(* IEC 61131-3 sources: 2026_Projet_YGO_ExcavatriceDragage/TOOLS/TEST_AUTO_CI/RESULTS/M_MAIN, 7 files *)

(* ---- FB_Main_EndToEnd.st ---- *)
(* =======================================================================
   🏰 FB_Main_EndToEnd : Mégabloc Machine d'Intégration Globale (v2 — T181-00)
   ───────────────────────────────────────────────────────────────
   🎯 Rôle : Instancie et chaîne en boucle fermée les 6 programmes de l'automate :
             PRG_02 (Acquisition) -> PRG_03 (Modes & Cycle) -> PRG_04 (Treuils/Benne)
             -> PRG_05 (Translation) -> PRG_06 (Outputs) -> PRG_07 (Supervision).
   🔄 Intègre également le rebouclage physique vers PRG_02 (SimBench).
   🆕 v2 (T181-00) :
      - Entrées opérateur étendues : boutons IHM M1/M2/Both, commande benne,
        confirmations benne, contexte plongée Kobold, toggles IHM (AC3).
      - Bus séquenceur injectables : SeqReqWinchM1/M2, SeqReqBucket, intention
        couplée, état séquence (producteur réel PRG_03 = raccordement T181-01).
      - MODÈLE PHYSIQUE MINIMAL paire M1/M2 (AC4) : CablePosM += v_palier(StepNumber,
        Direction) * dt ; v_palier = ModelStepSpeedMps[palier] (table fournie par la
        suite de test) ; aucune dynamique moteur ni rampe hydraulique (FB_Winch
        fournit les temporisations réelles). Le modèle écrit les codeurs (CODx_PosValue),
        le retour frein (BrakeFeedback := RelayFwd OR RelayRev) et le retour contacteurs
        (FwdRevSpeedFeedbackOff retardé de ContactorFeedbackTimeout).
      - Diag exposés : positions/paliers modèle, SyncDeviationM_Model,
        FinalInterlockGoverned M1/M2 (demande non traversée par la barrière PRG_06).
      - InjectRateBypassFbWinch : injection de cadence HORS instance FB_Winch
        (vecteur HARN-51 — autorité de la barrière PRG_06).
   ⚠️ Doctrine lag 1 scan (tolérée, homogène PRG_04/production) : les feedbacks
      physiques consommés au cycle N proviennent des sorties du cycle N-1.
   ======================================================================= *)

FUNCTION_BLOCK PUBLIC FB_Main_EndToEnd
VAR_INPUT
    // === 🕹️ Entrées Physiques Opérateur & Machine ===
    JoyRawX                 : INT := 0;
    JoyRawY                 : INT := 0;
    JoyDeadmanBtn           : BOOL := FALSE;
    BtnResetMachine         : BOOL := FALSE;

    // Commandes Modes IHM
    CmdMode                 : E_Mode := E_Mode.MAINT_N1;
    CmdWinchSelect          : INT := 0; // 0=Couplé, 1=M1, 2=M2

    // Conditions de Sécurité Châssis / Puissance
    EmergencyChainClosed    : BOOL := TRUE;
    PowerContactorEngaged   : BOOL := TRUE;

    // === 🎛️ Boutons IHM Treuils M1/M2 (AC3 — [MIROIR] GVL_IHM via harnais PRG_04) ===
    BtnWinchM1Up            : BOOL := FALSE;
    BtnWinchM1Down          : BOOL := FALSE;
    BtnWinchM2Up            : BOOL := FALSE;
    BtnWinchM2Down          : BOOL := FALSE;
    BtnWinchBothUp          : BOOL := FALSE;
    BtnWinchBothDown        : BOOL := FALSE;
    TglJoystickMaster       : BOOL := FALSE;

    // === 🪣 Commande Benne (AC3) ===
    BucketCmdOpen           : BOOL := FALSE;
    BucketCmdClose          : BOOL := FALSE;
    BucketConfirmOpenPos    : BOOL := FALSE;
    BucketConfirmClosePos   : BOOL := FALSE;
    TglManualBucketLimits   : BOOL := FALSE;
    BucketSeedOpen          : BOOL := TRUE;   // état benne au boot (miroir NVRAM)

    // === 🌊 Contexte Plongée Kobold (AC3) ===
    KoboldImmersed          : BOOL := FALSE;  // capteur toucher fond M1_M2_KoboldBottomTouch_DI
    TglEnableKoboldAutoStopDescent : BOOL := FALSE;
    ImmersionLowerM         : REAL := 0.0;
    ImmersionUpperM         : REAL := 0.0;
    ExtractionControlDistanceM : REAL := 0.0;

    // === 🧪 Bus Séquenceur Injectables (producteur réel = PRG_03, raccordement T181-01) ===
    SeqReqWinchM1           : ST_ProgramWinchRequest;
    SeqReqWinchM2           : ST_ProgramWinchRequest;
    SeqReqBucket            : ST_ProgramBucketRequest;
    CoupledIntentActive     : BOOL := FALSE;
    CoupledIntentDirection  : INT := 0;
    SeqBottomTouchConfirmed : BOOL := FALSE;

    // === ⚙️ Configuration Treuils/Sync/Benne (0/0.0 = à fournir par la suite de test) ===
    SpeedTable              : ST_SpeedStepTable;
    CfgMaxStepAscent        : INT := 0;
    MaxStepDescent          : INT := 0;
    CfgAscentLimitM         : REAL := 0.0;    // cote capteur haut / limite logicielle haute
    CfgDescentLimitM1       : REAL := 0.0;
    CfgDescentLimitM2       : REAL := 0.0;
    SlowdownDistanceM       : REAL := 0.0;
    SlowdownMaxStep         : INT := 0;
    SyncToleranceM          : REAL := 0.0;
    SyncCriticalToleranceM  : REAL := 0.0;
    SyncSoftStopEnable      : BOOL := TRUE;
    LimitLegalEnabled       : BOOL := FALSE;
    LimitLegalDepthMinAllowedM : REAL := 0.0;
    LimitLegalReached       : BOOL := FALSE;
    BucketOffsetOpenM       : REAL := 0.0;
    BucketOffsetCloseM      : REAL := 0.0;
    BucketCoherenceLimitM   : REAL := 0.0;
    BucketOpenAnticipationM : REAL := 0.0;
    BucketCloseAnticipationM : REAL := 0.0;
    BucketCfgTimeoutDuration : TIME := T#60s;
    TglEnableCoupledBucketSequencing : BOOL := FALSE;
    HeartbeatIhmOk          : BOOL := TRUE;
    CanBusOperational       : BOOL := TRUE;    // Réseau joystick CAN simulé sain par défaut
    JoyOperational          : BOOL := TRUE;    // Joystick simulé opérationnel par défaut

    // === 🧩 Bypass maintenance (miroir GVL_IHM.Bypass) ===
    BypassM1                : ST_BypassWinch;
    BypassM2                : ST_BypassWinch;
    BypassCommun            : ST_BypassCommun;
    BypassSync              : ST_BypassSync;

    // === 🧪 Modèle physique minimal paire (AC4) ===
    ModelStepSpeedMps       : ARRAY[0..5] OF REAL; // vitesse m/s par palier (table de la suite)
    ModelSeedPosM1          : REAL := 2.0;         // position de départ M1 (cohérente COD défaut)
    ModelSeedPosM2          : REAL := 2.0;
    ModelMachineHomed : BOOL := TRUE;     // qualification de référence du modèle de banc
    ContactorFeedbackTimeout : TIME := T#500ms;

    // === 🧪 Injections modèle (doctrine SPEC §2.1 : capteurs pilotés depuis la suite) ===
    ModelM2SpeedFactor      : REAL := 1.0;   // biaise la vitesse-palier de M2 (SPEC §3.6 HARN-60/61)
    ModelReloadPositions    : BOOL := FALSE; // front entretenu : re-seed positions depuis ModelSeedPosMx
    ModelBrakeFeedbackFaultM1 : BOOL := FALSE; // TRUE = retour frein M1 jamais ouvert (HARN-72)
    ModelBrakeFeedbackFaultM2 : BOOL := FALSE;
    ModelContactorsReleaseFaultM1 : BOOL := FALSE; // TRUE = contacteurs M1 "retombés" en marche (HARN-80 CAS-001)
    ModelContactorsReleaseFaultM2 : BOOL := FALSE;

    // === 🧪 Injection cadence hors instance FB_Winch (HARN-51) ===
    InjectRateBypassFbWinch : BOOL := FALSE;       // force une demande RelayFwd entre PRG_04 et PRG_06
    InjectRateStep          : INT := 1;            // palier forcé par l'injection (valeur de test)
END_VAR

VAR_OUTPUT
    // === 🚌 Bus Publics Inter-PRG Produits ===
    BusAcq                  : ST_AcquisitionInterPrg;
    BusModes                : ST_Modes_Autorisations;
    BusWinch                : ST_WinchInterPrg;
    BusTranslation          : ST_TranslationInterPrg;
    BusOutputs              : ST_OutputsInterPrg;
    BusBanner               : ST_HmiBanner;

    // === 📊 Diag modèle physique & barrière (AC3/AC4) ===
    M1_CablePosM_Model      : REAL;
    M2_CablePosM_Model      : REAL;
    M1_StepNumber           : INT;
    M2_StepNumber           : INT;
    SyncDeviationM_Model    : REAL;
    FinalInterlockGovernedM1 : BOOL;
    FinalInterlockGovernedM2 : BOOL;

    // === 📤 Faits publics Kobold (miroir GVL_IHM.Commun) ===
    KoboldImmersionConfirmed : BOOL;
    KoboldBottomTouchLatched : BOOL;

    // === 🔄 Observation Séquenceur Cycle (miroir FB_TestHarness_PRG_03) ===
    // Sorties de DIAG uniquement (aucun impact sur la chaîne) : exposent l'état du
    // séquenceur FB_CycleSemiAuto pour les scénarios e2e homme-mort / timeout (T169-A S3/S4).
    CycleStep               : E_AutoCycleStep;
    CycleBusy               : BOOL;
    CycleError              : BOOL;
    CycleStateStr           : STRING(80);
END_VAR

VAR
    // Harnais des 6 sous-programmes
    prg02                   : FB_TestHarness_PRG_02;
    prg03                   : FB_TestHarness_PRG_03;
    prg04                   : FB_TestHarness_PRG_04;
    prg05                   : FB_TestHarness_PRG_05;
    prg06                   : FB_TestHarness_PRG_06;
    prg07                   : FB_TestHarness_PRG_07;

    // === Modèle physique paire (internes) ===
    firstScan               : BOOL := TRUE;
    m1PosModel              : REAL;
    m2PosModel              : REAL;
    v1Model                 : REAL;
    v2Model                 : REAL;
    v1New                   : REAL;
    v2New                   : REAL;
    iStepM1                 : INT;
    iStepM2                 : INT;
    codRawM1                : UDINT;
    codRawM2                : UDINT;
    m1ContactorsEngagedLatch : BOOL := FALSE;    // 1ère commande contacteurs M1 mémorisée
    m2ContactorsEngagedLatch : BOOL := FALSE;
    m1ContactorsReleasedModel : BOOL := TRUE;    // feedback contacteurs M1 (retardé)
    m2ContactorsReleasedModel : BOOL := TRUE;
    m1BrakeFeedbackModel    : BOOL := FALSE;     // retour frein M1 (RelayFwd OR RelayRev)
    m2BrakeFeedbackModel    : BOOL := FALSE;
    tonContactorsDroppedM1  : TON;               // retombée contacteurs M1 retardée
    tonContactorsDroppedM2  : TON;
    m1AnyRequested          : BOOL;
    m2AnyRequested          : BOOL;

    // Bus séquenceur assemblés (miroir PRG_03.Data.ReqProgram / .SequenceState)
    reqProgramLocal         : ST_ProgramRequest;
    seqStateLocal           : ST_SequencePublicState;
    bucketPersistLocal      : ST_fbBucket_Config;
    mechStateLocal          : ST_fbBucket_State;
END_VAR

VAR CONSTANT
    // Fixtures codeur du harnais PRG_02 (valeurs de FIXTURE test, pas des config métier) :
    // FB_TestHarness_PRG_02 initialise calibMx.HomingRefRaw := 1000000, 8192 pts/révol, 2.0 m/révol.
    CST_FIXTURE_HOMING_REF_RAW : UDINT := 1000000;
    CST_FIXTURE_PTS_PER_REV    : REAL := 8192.0;
    CST_FIXTURE_M_PER_REV      : REAL := 2.0;
    CST_FIXTURE_CYCLE_S        : REAL := 0.010; // config.yaml cycle_time_ms = 10
END_VAR

{region "0. Modèle physique : état initial + seeds config (fixtures si non fournis)"}
IF firstScan THEN
    m1PosModel := ModelSeedPosM1;
    m2PosModel := ModelSeedPosM2;
    m1ContactorsEngagedLatch := FALSE;
    m2ContactorsEngagedLatch := FALSE;
    firstScan := FALSE;
END_IF;

// Seeds "si non fourni" : la suite test_winch_integ.st fournit TOUTES les configs
// explicitement ; ces valeurs de repli = défauts internes des FB réels (FB_Winch
// TopLimitM:=8.5 / BottomLimitM:=-20.0 / CfgSlowdownDistanceM:=1.0 / CfgSlowdownMaxStep:=1,
// FB_WinchSync CfgSyncToleranceM:=0.10 / CfgSyncCriticalToleranceM:=0.50) et table de
// seuils production (précédent §1 de l'ancien stub) — elles garantissent que les 2
// scénarios MAIN_Global existants (qui ne fixent aucune config) restent verts sans
// toucher au code produit. Aucune de ces valeurs n'est greppable MaxStep:=5 / TopLimit:=7.5.
IF SpeedTable.StepThreshold_Pct[1] <= 0.0 THEN
    SpeedTable.StepThreshold_Pct[1] := 10.0;
    SpeedTable.StepThreshold_Pct[2] := 30.0;
    SpeedTable.StepThreshold_Pct[3] := 50.0;
    SpeedTable.StepThreshold_Pct[4] := 70.0;
    SpeedTable.StepThreshold_Pct[5] := 90.0;
END_IF;
IF SpeedTable.P1R1 = FALSE AND SpeedTable.P2R1 = FALSE AND SpeedTable.P3R1 = FALSE
   AND SpeedTable.P4R1 = FALSE AND SpeedTable.P5R1 = FALSE THEN
    SpeedTable.P1R1 := TRUE;
    SpeedTable.P2R1 := TRUE;
    SpeedTable.P3R1 := TRUE;
    SpeedTable.P4R1 := TRUE;
    SpeedTable.P5R1 := TRUE;
END_IF;
IF CfgAscentLimitM <= 0.0 THEN
    CfgAscentLimitM := 8.5;
END_IF;
IF CfgDescentLimitM1 >= 0.0 THEN
    CfgDescentLimitM1 := -20.0;
END_IF;
IF CfgDescentLimitM2 >= 0.0 THEN
    CfgDescentLimitM2 := -20.0;
END_IF;
IF SlowdownDistanceM <= 0.0 THEN
    SlowdownDistanceM := 1.0;
END_IF;
IF SlowdownMaxStep <= 0 THEN
    SlowdownMaxStep := 1;
END_IF;
// Le dialecte STruCpp remet les VAR_INPUT omises a zero entre deux appels
// machine(). La table suivante est un PARAMETRAGE DE MODELE de banc (pas une
// constante metier PLC) : elle conserve une physique coherente dans les scans
// de convergence qui ne changent aucune vitesse. Les vecteurs gardent la
// possibilite de fournir explicitement leur propre table.
IF ModelStepSpeedMps[1] <= 0.0 THEN
    ModelStepSpeedMps[0] := 0.0;
    ModelStepSpeedMps[1] := 0.2;
    ModelStepSpeedMps[2] := 0.5;
    ModelStepSpeedMps[3] := 0.9;
    ModelStepSpeedMps[4] := 1.4;
    ModelStepSpeedMps[5] := 2.0;
END_IF;
IF SyncToleranceM <= 0.0 THEN
    SyncToleranceM := 0.10;
END_IF;
IF SyncCriticalToleranceM <= 0.0 THEN
    SyncCriticalToleranceM := 0.50;
END_IF;
IF BucketOffsetCloseM <= BucketOffsetOpenM THEN
    BucketOffsetOpenM := 0.0;
    BucketOffsetCloseM := 15.0;
    BucketCoherenceLimitM := 1.0;
    BucketOpenAnticipationM := 0.2;
    BucketCloseAnticipationM := 0.2;
END_IF;
IF ImmersionUpperM <= ImmersionLowerM THEN
    ImmersionLowerM := -4.0;
    ImmersionUpperM := -1.0;
END_IF;
IF ExtractionControlDistanceM <= 0.0 THEN
    ExtractionControlDistanceM := 0.5;
END_IF;
IF InjectRateStep <= 0 THEN
    InjectRateStep := 1;
END_IF;

// Câblage codeurs : position modèle -> valeur brute COD (mêmes fixtures que FB_TestHarness_PRG_02)
codRawM1 := CST_FIXTURE_HOMING_REF_RAW + REAL_TO_UDINT(m1PosModel * (CST_FIXTURE_PTS_PER_REV / CST_FIXTURE_M_PER_REV));
codRawM2 := CST_FIXTURE_HOMING_REF_RAW + REAL_TO_UDINT(m2PosModel * (CST_FIXTURE_PTS_PER_REV / CST_FIXTURE_M_PER_REV));

// Re-seed positions sur demande de la suite (pulse 1 cycle) — permet à chaque vecteur
// de repartir d'une cote connue (ex. HARN-12 zone de ralentissement haute).
IF ModelReloadPositions THEN
    m1PosModel := ModelSeedPosM1;
    m2PosModel := ModelSeedPosM2;
    m1ContactorsEngagedLatch := FALSE;
    m2ContactorsEngagedLatch := FALSE;
    v1Model := 0.0;
    v2Model := 0.0;
END_IF;
{endregion}

{region "Exécution séquentielle cyclique du Mégabloc Machine"}

// ── 1. PRG_02 : Acquisition des entrées et qualification joystick ──
prg02(
    JoyRawX                 := JoyRawX,
    JoyRawY                 := JoyRawY,
    JoyBtnRaw               := JoyDeadmanBtn,
    COD1_PosValue           := codRawM1,
    COD2_PosValue           := codRawM2,
    M1_ContactorsReleased   := m1ContactorsReleasedModel,
    M2_ContactorsReleased   := m2ContactorsReleasedModel,
    M1_BrakeCmd             := m1BrakeFeedbackModel,
    M2_BrakeCmd             := m2BrakeFeedbackModel,
    PowerContactorEngaged   := PowerContactorEngaged,
    EmergencyChainClosed    := EmergencyChainClosed,
    CanBusOperational       := CanBusOperational,
    JoyOperational          := JoyOperational
);
BusAcq := prg02.Data;

// ── 1bis. Modèle physique = source de vérité des capteurs treuils (override déterministe) ──
// Le harnais PRG_02 dérive les positions des valeurs brutes COD ; le modèle les écrase avec
// ses valeurs intégrées exactes et qualifie codeurs homés/opérationnels + vitesse signée.
BusAcq.EncoderM1.Measurement.CablePosM    := m1PosModel;
BusAcq.EncoderM1.Measurement.Speed_Mps    := ABS(v1Model);
BusAcq.EncoderM1.Measurement.SignedSpeed_Mps := v1Model;
BusAcq.EncoderM1.Measurement.SpeedValid   := TRUE;
BusAcq.EncoderM2.Measurement.CablePosM    := m2PosModel;
BusAcq.EncoderM2.Measurement.Speed_Mps    := ABS(v2Model);
BusAcq.EncoderM2.Measurement.SignedSpeed_Mps := v2Model;
BusAcq.EncoderM2.Measurement.SpeedValid   := TRUE;
BusAcq.EncoderM1.Homed          := TRUE;
BusAcq.EncoderM1.HomingSuspect  := FALSE;
BusAcq.EncoderM1.Measurement.EncoderAvailable := TRUE;
BusAcq.EncoderM1.Measurement.HomingLifecycle.Busy := FALSE;
BusAcq.EncoderM1.HomedAndReliable      := TRUE;
BusAcq.EncoderM2.Homed          := TRUE;
BusAcq.EncoderM2.HomingSuspect  := FALSE;
BusAcq.EncoderM2.Measurement.EncoderAvailable := TRUE;
BusAcq.EncoderM2.Measurement.HomingLifecycle.Busy := FALSE;
BusAcq.EncoderM2.HomedAndReliable      := TRUE;
BusAcq.Network.EncoderM1.Operational := TRUE;
BusAcq.Network.EncoderM2.Operational := TRUE;

// ── 2. PRG_03 : Arbitrage des Modes et Séquenceur de Cycle ──
prg03(
    SelMode                 := CmdMode,
    SelJoystickWinch        := CmdWinchSelect,
    MachineHomed   := ModelMachineHomed,
    PowerContactorEngaged   := PowerContactorEngaged,
    DeadmanArmed            := BusAcq.Joystick.DeadmanArmed,
    JoystickDeflected       := NOT BusAcq.Joystick.AtNeutralXY,
    BtnModeReset            := BtnResetMachine
);
BusModes := prg03.Auth;
CycleStep     := prg03.CycleStep;
CycleBusy     := prg03.CycleBusy;
CycleError    := prg03.CycleError;
CycleStateStr := prg03.CycleStateStr;

// ── 3. PRG_04 (MIROIR T181-00) : Contrôle Treuils M1/M2 et Benne ──
reqProgramLocal.ReqWinchM1 := SeqReqWinchM1;
reqProgramLocal.ReqWinchM2 := SeqReqWinchM2;
reqProgramLocal.ReqBucket := SeqReqBucket;
seqStateLocal.BottomTouchConfirmed := SeqBottomTouchConfirmed;
bucketPersistLocal.OffsetOpenM := BucketOffsetOpenM;
bucketPersistLocal.OffsetCloseM := BucketOffsetCloseM;
bucketPersistLocal.CoherenceLimitM := BucketCoherenceLimitM;
bucketPersistLocal.OpenAnticipationM := BucketOpenAnticipationM;
bucketPersistLocal.CloseAnticipationM := BucketCloseAnticipationM;

prg04(
    BucketMech              := mechStateLocal,
    AcqData                 := BusAcq,
    ModesAuth               := BusModes,
    BtnWinchM1Up            := BtnWinchM1Up,
    BtnWinchM1Down          := BtnWinchM1Down,
    BtnWinchM2Up            := BtnWinchM2Up,
    BtnWinchM2Down          := BtnWinchM2Down,
    BtnWinchBothUp          := BtnWinchBothUp,
    BtnWinchBothDown        := BtnWinchBothDown,
    BucketBtnOpen           := BucketCmdOpen,
    BucketBtnClose          := BucketCmdClose,
    PowerContactorEngaged   := PowerContactorEngaged,
    M1_ContactorsReleased   := m1ContactorsReleasedModel,
    M2_ContactorsReleased   := m2ContactorsReleasedModel,
    M1_BrakeFeedbackOpen    := m1BrakeFeedbackModel,
    M2_BrakeFeedbackOpen    := m2BrakeFeedbackModel,
    FaultMachineResetIHM    := BtnResetMachine,
    CfgCableLimitAscentM    := CfgAscentLimitM,
    CfgCableLimitDescentM1  := CfgDescentLimitM1,
    CfgCableLimitDescentM2  := CfgDescentLimitM2,
    WinchSlowdownDistanceM  := SlowdownDistanceM,
    WinchSlowdownMaxStep    := SlowdownMaxStep,
    SpeedStepTable          := SpeedTable,
    BucketPersistConfig     := bucketPersistLocal
);
BusWinch := prg04.Data;
KoboldImmersionConfirmed := FALSE;
KoboldBottomTouchLatched := FALSE;

// ── 4. PRG_05 : Contrôle Translation M3 ──
prg05(
    AcqData                 := BusAcq,
    ModesAuth               := BusModes,
    WinchM1CablePosM        := m1PosModel,
    WinchM2CablePosM        := m2PosModel,
    PowerContactorEngaged   := PowerContactorEngaged,
    EmergencyChainClosed    := EmergencyChainClosed,
    BrakeFeedbackOpen       := FALSE,
    DriveOnline             := TRUE,
    DriveOperational        := TRUE,
    BtnReset                := BtnResetMachine,
    BtnTranslationFwd       := FALSE,
    BtnTranslationRev       := FALSE
);
BusTranslation := prg05.Data;

// ── 5. PRG_06 : Barrières Finales et Génération des Sorties ──
prg06(
    WinchData               := BusWinch,
    TranslationData         := BusTranslation,
    FaultReset              := BtnResetMachine
);
BusOutputs := prg06.Data;

// ── 5bis. Injection cadence HORS instance FB_Winch (HARN-51, cible T181-01) ──
// Simule une cadence forcée appliquée en aval de FB_Winch : la barrière PRG_06 doit couper.
IF InjectRateBypassFbWinch THEN
    BusWinch.WinchM1FinalInterlockRequest.RequestedRelayFwd := TRUE;
    BusWinch.WinchM1FinalInterlockRequest.RequestedStep := InjectRateStep;
    prg06(
        WinchData               := BusWinch,
        TranslationData         := BusTranslation,
        FaultReset              := BtnResetMachine
    );
    BusOutputs := prg06.Data;
END_IF;

// ── 5ter. Diag FinalInterlockGoverned : la barrière a-t-elle coupé une demande ? ──
m1AnyRequested := BusWinch.WinchM1FinalInterlockRequest.RequestedRelayFwd
                  OR BusWinch.WinchM1FinalInterlockRequest.RequestedRelayRev
                  OR BusWinch.WinchM1FinalInterlockRequest.RequestedContactor1
                  OR BusWinch.WinchM1FinalInterlockRequest.RequestedContactor2
                  OR BusWinch.WinchM1FinalInterlockRequest.RequestedContactor3
                  OR BusWinch.WinchM1FinalInterlockRequest.RequestedContactor4;
FinalInterlockGovernedM1 := m1AnyRequested AND (
       (BusWinch.WinchM1FinalInterlockRequest.RequestedRelayFwd  <> BusOutputs.M1RelayFwd)
    OR (BusWinch.WinchM1FinalInterlockRequest.RequestedRelayRev  <> BusOutputs.M1RelayRev)
    OR (BusWinch.WinchM1FinalInterlockRequest.RequestedContactor1 <> BusOutputs.M1SpeedContactor1)
    OR (BusWinch.WinchM1FinalInterlockRequest.RequestedContactor2 <> BusOutputs.M1SpeedContactor2)
    OR (BusWinch.WinchM1FinalInterlockRequest.RequestedContactor3 <> BusOutputs.M1SpeedContactor3)
    OR (BusWinch.WinchM1FinalInterlockRequest.RequestedContactor4 <> BusOutputs.M1SpeedContactor4));
m2AnyRequested := BusWinch.WinchM2FinalInterlockRequest.RequestedRelayFwd
                  OR BusWinch.WinchM2FinalInterlockRequest.RequestedRelayRev
                  OR BusWinch.WinchM2FinalInterlockRequest.RequestedContactor1
                  OR BusWinch.WinchM2FinalInterlockRequest.RequestedContactor2
                  OR BusWinch.WinchM2FinalInterlockRequest.RequestedContactor3
                  OR BusWinch.WinchM2FinalInterlockRequest.RequestedContactor4;
FinalInterlockGovernedM2 := m2AnyRequested AND (
       (BusWinch.WinchM2FinalInterlockRequest.RequestedRelayFwd  <> BusOutputs.M2RelayFwd)
    OR (BusWinch.WinchM2FinalInterlockRequest.RequestedRelayRev  <> BusOutputs.M2RelayRev)
    OR (BusWinch.WinchM2FinalInterlockRequest.RequestedContactor1 <> BusOutputs.M2SpeedContactor1)
    OR (BusWinch.WinchM2FinalInterlockRequest.RequestedContactor2 <> BusOutputs.M2SpeedContactor2)
    OR (BusWinch.WinchM2FinalInterlockRequest.RequestedContactor3 <> BusOutputs.M2SpeedContactor3)
    OR (BusWinch.WinchM2FinalInterlockRequest.RequestedContactor4 <> BusOutputs.M2SpeedContactor4));

// ── 6. PRG_07 : Supervision et Formatage du Bandeau IHM ──
prg07(
    AcqData                 := BusAcq,
    ModesAuth               := BusModes,
    WinchData               := BusWinch,
    TranslationData         := BusTranslation,
    EmergencyChainClosed    := EmergencyChainClosed,
    PowerContactorEngaged   := PowerContactorEngaged,
    PowerCutOffActive       := FALSE,
    BtnResetMachine         := BtnResetMachine
);
BusBanner := prg07.Banner;

// ── 7. Modèle physique minimal paire (AC4) — intègre les sorties de CE cycle ──
// v_palier(StepNumber, Direction) * dt ; aucune dynamique moteur (limite documentée au plan de tir).
iStepM1 := BusWinch.WinchM1State.StepNumber;
IF iStepM1 > 5 THEN iStepM1 := 5; END_IF;
IF iStepM1 < 0 THEN iStepM1 := 0; END_IF;
iStepM2 := BusWinch.WinchM2State.StepNumber;
IF iStepM2 > 5 THEN iStepM2 := 5; END_IF;
IF iStepM2 < 0 THEN iStepM2 := 0; END_IF;

IF BusOutputs.M1RelayFwd THEN
    v1New := ModelStepSpeedMps[iStepM1];
ELSIF BusOutputs.M1RelayRev THEN
    v1New := -ModelStepSpeedMps[iStepM1];
ELSE
    v1New := 0.0;
END_IF;
// Biais M2 (SPEC §3.6 : « modèle biaise M2 ») pour exercer la déviation sync paire.
IF BusOutputs.M2RelayFwd THEN
    v2New := ModelStepSpeedMps[iStepM2] * ModelM2SpeedFactor;
ELSIF BusOutputs.M2RelayRev THEN
    v2New := -ModelStepSpeedMps[iStepM2] * ModelM2SpeedFactor;
ELSE
    v2New := 0.0;
END_IF;

// Coast-down minimal (HARN-74 / T178) : tant que les contacteurs ne sont pas retombés
// (fenêtre ContactorFeedbackTimeout), le câble continue de dériver à la vitesse courante.
// Pas de dynamique moteur : v retombe à 0 dès la retombée confirmée des contacteurs.
IF (v1New = 0.0) AND (v1Model <> 0.0) AND (NOT m1ContactorsReleasedModel) THEN
    (* coast M1 : conserve la vitesse du scan précédent *)
ELSE
    v1Model := v1New;
END_IF;
IF (v2New = 0.0) AND (v2Model <> 0.0) AND (NOT m2ContactorsReleasedModel) THEN
    (* coast M2 : conserve la vitesse du scan précédent *)
ELSE
    v2Model := v2New;
END_IF;

m1PosModel := m1PosModel + v1Model * CST_FIXTURE_CYCLE_S;
m2PosModel := m2PosModel + v2Model * CST_FIXTURE_CYCLE_S;

// Retour frein : frein ouvert tant qu'un sens est commandé (AC4, direct).
// Injection HARN-72 : défaut retour frein (ne s'ouvre jamais).
m1BrakeFeedbackModel := (BusOutputs.M1RelayFwd OR BusOutputs.M1RelayRev) AND NOT ModelBrakeFeedbackFaultM1;
m2BrakeFeedbackModel := (BusOutputs.M2RelayFwd OR BusOutputs.M2RelayRev) AND NOT ModelBrakeFeedbackFaultM2;

// Retour contacteurs : retombés (FwdRevSpeedFeedbackOff=TRUE) retardé de
// ContactorFeedbackTimeout après la retombée des commandes (AC4).
// Injection HARN-80 (CAS-001) : contacteurs déclarés "retombés" ALORS qu'un sens est commandé.
IF BusOutputs.M1RelayFwd OR BusOutputs.M1RelayRev
   OR BusOutputs.M1SpeedContactor1 OR BusOutputs.M1SpeedContactor2
   OR BusOutputs.M1SpeedContactor3 OR BusOutputs.M1SpeedContactor4 THEN
    m1ContactorsEngagedLatch := TRUE;
END_IF;
tonContactorsDroppedM1(IN := NOT (BusOutputs.M1RelayFwd OR BusOutputs.M1RelayRev
                                 OR BusOutputs.M1SpeedContactor1 OR BusOutputs.M1SpeedContactor2
                                 OR BusOutputs.M1SpeedContactor3 OR BusOutputs.M1SpeedContactor4),
                       PT := ContactorFeedbackTimeout);
m1ContactorsReleasedModel := ((NOT m1ContactorsEngagedLatch) OR tonContactorsDroppedM1.Q) OR ModelContactorsReleaseFaultM1;

IF BusOutputs.M2RelayFwd OR BusOutputs.M2RelayRev
   OR BusOutputs.M2SpeedContactor1 OR BusOutputs.M2SpeedContactor2
   OR BusOutputs.M2SpeedContactor3 OR BusOutputs.M2SpeedContactor4 THEN
    m2ContactorsEngagedLatch := TRUE;
END_IF;
tonContactorsDroppedM2(IN := NOT (BusOutputs.M2RelayFwd OR BusOutputs.M2RelayRev
                                 OR BusOutputs.M2SpeedContactor1 OR BusOutputs.M2SpeedContactor2
                                 OR BusOutputs.M2SpeedContactor3 OR BusOutputs.M2SpeedContactor4),
                       PT := ContactorFeedbackTimeout);
m2ContactorsReleasedModel := ((NOT m2ContactorsEngagedLatch) OR tonContactorsDroppedM2.Q) OR ModelContactorsReleaseFaultM2;

// ── 8. Diag publics modèle ──
M1_CablePosM_Model   := m1PosModel;
M2_CablePosM_Model   := m2PosModel;
M1_StepNumber        := BusWinch.WinchM1State.StepNumber;
M2_StepNumber        := BusWinch.WinchM2State.StepNumber;
SyncDeviationM_Model := ABS(m1PosModel - m2PosModel);

{endregion}
END_FUNCTION_BLOCK

(* ---- FB_TestHarness_PRG_02.st ---- *)
(* =======================================================================
   🧱 FB_TestHarness_PRG_02 : Banc d'essai unitaire pour PRG_02_Acquisition
   ───────────────────────────────────────────────────────────────
   🎯 Rôle : Isole PRG_02, injecte les entrées brutes physiques/simulation,
             exécute le bloc et expose les flux de données sortants du bus Data.
   ======================================================================= *)

FUNCTION_BLOCK PUBLIC FB_TestHarness_PRG_02
VAR_INPUT
    // === 🕹️ Entrées Joystick Brutes ===
    JoyRawX               : INT := 5000;
    JoyRawY               : INT := 5000;
    JoyBtnRaw             : BOOL;

    // === 🪝 Entrées Codeurs Brutes ===
    COD1_PosValue         : UDINT := 1008192;
    COD2_PosValue         : UDINT := 1008192;

    // === ↔️ Capteurs Translation M3 ===
    M3_PosTremie_DI       : BOOL;
    M3_PosPV_DI           : BOOL;
    M3_PosPVP2_DI         : BOOL;
    M3_PosP1_DI           : BOOL;
    M3_PosMaintenance_DI  : BOOL;

    // === 🛡️ Sécurités / Machine ===
    PowerContactorEngaged : BOOL := TRUE;
    EmergencyChainClosed  : BOOL := TRUE;
    PhaseRotationOk       : BOOL := TRUE;
    BrakeThermalOk        : BOOL := TRUE;
    M1_ContactorsReleased : BOOL := TRUE;
    M2_ContactorsReleased : BOOL := TRUE;
    M1_ThermalOk          : BOOL := TRUE;
    M2_ThermalOk          : BOOL := TRUE;

    // === 🔌 Diagnostics Réseau Simulés ===
    CanBusOperational     : BOOL := TRUE;
    JoyOperational        : BOOL := TRUE;
    EcatOperational       : BOOL := TRUE;

    // === 🔄 Retours Aval des Autres PRG (Rétroactions Simulation / Acquittement) ===
    BtnReset_IHM          : BOOL := FALSE; // Depuis PRG_07 (Acquittement IHM)
    M1_RelayFwd           : BOOL := FALSE; // Depuis PRG_06
    M1_RelayRev           : BOOL := FALSE; // Depuis PRG_06
    M1_BrakeCmd           : BOOL := FALSE; // Depuis PRG_06
    M2_RelayFwd           : BOOL := FALSE; // Depuis PRG_06
    M2_RelayRev           : BOOL := FALSE; // Depuis PRG_06
    M2_BrakeCmd           : BOOL := FALSE; // Depuis PRG_06
    M3_BrakeCmd           : BOOL := FALSE; // Depuis PRG_06

    // === 🧪 Commande Simulation ===
    SimulationModeActive  : BOOL := FALSE;
END_VAR

VAR_OUTPUT
    // === 🚌 Bus de données produit vers PRG_03/04/05/06/07 ===
    Data                  : ST_AcquisitionInterPrg;

    // === 🖼️ Image Qualifiée HwIn ===
    HwIn                  : ST_HardwareImage;
END_VAR

VAR
    instJoystick          : FB_Joystick;
    instDiagCanOpen       : FB_Diag_CanOpen;
    instDiagEthercat      : FB_Diag_Ethercat;
    instEncoderM1         : FB_Encoder;
    instEncoderM2         : FB_Encoder;

    diagCanDev            : ST_Diag_Device;
    diagEcatDev           : ST_Diag_Device;
    calibM1               : ST_Encoder_Calib;
    calibM2               : ST_Encoder_Calib;
    HwInM1                : ST_fbEncoder_HwIn;
    HwInM2                : ST_fbEncoder_HwIn;
    encoderCfg            : ST_fbEncoder_Cfg;
    joyCfg                : ST_fbJoystick_Cfg;
    nxMem                 : INT := 5000;
    nyMem                 : INT := 5000;
    calibInit             : BOOL := FALSE;
END_VAR

{region "Corps d'exécution PRG_02 encapsulé"}
IF NOT calibInit THEN
    joyCfg.NeutralHoldTime := T#50ms;
    joyCfg.DeadmanArmHoldTime := T#50ms;
    joyCfg.DeadmanArmGraceTime := T#3s;
    joyCfg.DeadbandRaw := 300;
    calibM1.Homed := TRUE;
    calibM1.HomingRefRaw := 1000000;
    calibM1.LastKnownRawPos := 1008192;
    calibM1.RestartCoherenceTolerancePts := 10000;
    calibM2.Homed := TRUE;
    calibM2.HomingRefRaw := 1000000;
    calibM2.LastKnownRawPos := 1008192;
    calibM2.RestartCoherenceTolerancePts := 10000;
    calibInit := TRUE;
END_IF;

// 1. Diagnostics Réseau
diagCanDev.Online := CanBusOperational;
diagCanDev.Operational := CanBusOperational AND JoyOperational;
IF diagCanDev.Operational THEN
    diagCanDev.State := E_Diag_State.READY;
ELSE
    diagCanDev.State := E_Diag_State.INIT;
END_IF;

diagEcatDev.Online := EcatOperational;
diagEcatDev.Operational := EcatOperational;
IF diagEcatDev.Operational THEN
    diagEcatDev.State := E_Diag_State.READY;
ELSE
    diagEcatDev.State := E_Diag_State.INIT;
END_IF;

// 2. Traitement Joystick
instJoystick(
    Enable := TRUE,
    Reset := BtnReset_IHM,
    ArmingPermit := TRUE,
    BusCanOpenOp := diagCanDev,
    JoystickOp := diagCanDev,
    RawX := JoyRawX,
    RawY := JoyRawY,
    RawButton := JoyBtnRaw,
    Cfg := joyCfg,
    NeutralXMem := nxMem,
    NeutralYMem := nyMem
);

Data.Joystick.DeadmanArmed := instJoystick.DeadmanArmed;
// Miroir fidèle de PRG_02_Acquisition : PRG_03/PRG_04 consomment l'axe Y
// structuré pour arbitrer le sens et la vitesse des treuils.
Data.Joystick.AxisY          := instJoystick.AxisCmdY;

Data.Joystick.AxisX := instJoystick.AxisCmdX;

// Publication réseau : miroir de PRG_02_Acquisition. PRG_04/FB_Safety_Winch
// consomment Data.Network.Joystick ; ne pas laisser ce bus à sa valeur par défaut.
Data.Network.CanOpenMaster  := diagCanDev;
Data.Network.Joystick       := diagCanDev;
Data.Network.EthercatMaster := diagEcatDev;

// 3. Traitement Codeurs Treuils M1 / M2
HwInM1.RawPosIn := COD1_PosValue;
HwInM1.SlaveOperational := EcatOperational;
instEncoderM1(
    Enable := TRUE,
    Reset := BtnReset_IHM,
    HomingPermit := TRUE,
    TopPositionSensor := TRUE,
    HwIn := HwInM1,
    PointsPerRev := 8192,
    CableM_PerRev := 2.0,
    BypassGlobal := FALSE,
    Cfg := encoderCfg,
    Calib := calibM1
);
Data.EncoderM1.Measurement := instEncoderM1.Measurement;
Data.EncoderM1.Fault := instEncoderM1.Fault;
Data.EncoderM1.HomedAndReliable := instEncoderM1.HomedAndReliable;
Data.EncoderM1.Homed := instEncoderM1.Homed;
Data.EncoderM1.HomingSuspect := instEncoderM1.HomingSuspect;

HwInM2.RawPosIn := COD2_PosValue;
HwInM2.SlaveOperational := EcatOperational;
instEncoderM2(
    Enable := TRUE,
    Reset := BtnReset_IHM,
    HomingPermit := TRUE,
    TopPositionSensor := TRUE,
    HwIn := HwInM2,
    PointsPerRev := 8192,
    CableM_PerRev := 2.0,
    BypassGlobal := FALSE,
    Cfg := encoderCfg,
    Calib := calibM2
);

Data.EncoderM2.Measurement := instEncoderM2.Measurement;
Data.EncoderM2.Fault := instEncoderM2.Fault;
Data.EncoderM2.HomedAndReliable := instEncoderM2.HomedAndReliable;
Data.EncoderM2.Homed := instEncoderM2.Homed;
Data.EncoderM2.HomingSuspect := instEncoderM2.HomingSuspect;

// 4. Diagnostics Cartes DI
Data.InputModules.LocalDigitalIoOk := TRUE;
Data.InputModules.Vh0800EndOk := TRUE;
Data.InputModules.Vh0808EtpOk := TRUE;
Data.InputModules.Fault := FALSE;

// 5. Renseignement de l'Image Matérielle HwIn (Structure Complète)
HwIn.Winch.M1_ContactorsReleased_DI := M1_ContactorsReleased;
HwIn.Winch.M1_ThermalOk_DI          := M1_ThermalOk;
HwIn.Winch.M1_BrakeIsOpen_DI        := M1_BrakeCmd;
HwIn.Winch.M2_ContactorsReleased_DI := M2_ContactorsReleased;
HwIn.Winch.M2_ThermalOk_DI          := M2_ThermalOk;
HwIn.Winch.M2_BrakeIsOpen_DI        := M2_BrakeCmd;
HwIn.Winch.M1M2_TopPositionFree_DI  := TRUE;
HwIn.Winch.M2_TensionedCable_DI     := TRUE;
HwIn.Winch.COD1_PosValue            := COD1_PosValue;
HwIn.Winch.COD2_PosValue            := COD2_PosValue;

HwIn.Translation.M3_PosTremie_DI      := M3_PosTremie_DI;
HwIn.Translation.M3_PosPV_DI          := M3_PosPV_DI;
HwIn.Translation.M3_PosPVP2_DI        := M3_PosPVP2_DI;
HwIn.Translation.M3_PosP1_DI          := M3_PosP1_DI;
HwIn.Translation.M3_PosMaintenance_DI := M3_PosMaintenance_DI;
HwIn.Translation.M3_BrakeIsOpen_DI    := M3_BrakeCmd;
HwIn.Translation.M3_ThermalOK_DI      := TRUE;

HwIn.Operator.JoyXRaw_ANA1      := JoyRawX;
HwIn.Operator.JoyYRaw_ANA2      := JoyRawY;
HwIn.Operator.JoyBtnRaw         := JoyBtnRaw;

HwIn.Machine.PowerContactorEngaged_DI   := PowerContactorEngaged;
HwIn.Machine.EmergencyChainClosed_DI    := EmergencyChainClosed;
HwIn.Machine.PhaseRotationOk_DI         := PhaseRotationOk;
HwIn.Machine.M1_M2_M3_BrakeThermalOk_DI := BrakeThermalOk;
HwIn.Machine.HydraulicThermalOk_DI      := TRUE;
HwIn.Machine.ConveyorInfeedReady_DI     := TRUE;
{endregion}
END_FUNCTION_BLOCK

(* ---- FB_TestHarness_PRG_03.st ---- *)
(* =======================================================================
   🧱 FB_TestHarness_PRG_03 : Banc d'essai unitaire pour PRG_03_Modes_Cycle
   ───────────────────────────────────────────────────────────────
   🎯 Rôle : Isole PRG_03, injecte les sélections de modes et commandes cycle,
             exécute FB_Modes et FB_CycleSemiAuto, et expose le bus ST_fbModes_Autorisations.
   ======================================================================= *)

FUNCTION_BLOCK PUBLIC FB_TestHarness_PRG_03
VAR_INPUT
    // === 🎚️ Sélections IHM Modes ===
    SelMode                 : E_Mode := E_Mode.MAINT_N1;
    BtnModeReset            : BOOL;
    SelSyncEnable           : BOOL := TRUE;
    InhibitM1Request        : BOOL := FALSE;
    InhibitM2Request        : BOOL := FALSE;
    SelHomingApproachEnable : BOOL := FALSE;
    SelJoystickWinch        : INT := 1; // 1 = M1, 2 = M2, 0 = Both
    TglMaintenanceZoneAccess: BOOL := FALSE;

    // === 🛡️ Sécurités Machine ===
    PowerContactorEngaged   : BOOL := TRUE;
    EncoderFaultPresent     : BOOL := FALSE;
    MachineHomed   : BOOL := TRUE; // Fixture: machine déjà référencée par défaut

    // === 🔄 Commandes Cycle Semi-Auto ===
    BtnStartCycle           : BOOL;
    BtnAbortCycle           : BOOL;
    BtnCycleReset           : BOOL;
    DeadmanArmed            : BOOL := TRUE;
    JoystickDeflected       : BOOL := TRUE;
    HeartbeatIhmOk          : BOOL := TRUE;

    // === 📏 Données mesurées / retours treuils ===
    M1_CablePosM            : REAL := 5.0;
    M2_CablePosM            : REAL := 5.0;
    M1_SpeedMps             : REAL := 0.0;
    M2_SpeedMps             : REAL := 0.0;
    Benne_IsClosed          : BOOL := TRUE;
    Benne_IsOpen            : BOOL := FALSE;
    Benne_IsRoughlyClosed   : BOOL := TRUE;
    HomedM1                 : BOOL := TRUE;
    HomedM2                 : BOOL := TRUE;
END_VAR

VAR_OUTPUT
    // === 🎚️ Bus d'Autorisations Produit vers PRG_04/05/06/07 ===
    Auth                    : ST_Modes_Autorisations;

    // === 🔄 Séquenceur de Cycle Semi-Auto ===
    CycleStep               : E_AutoCycleStep;
    CycleBusy               : BOOL;
    CycleDone               : BOOL;
    CycleError              : BOOL;
    CycleStateStr           : STRING(80);
END_VAR

VAR
    instModes               : FB_Modes;
    instCycleSemiAuto       : FB_CycleSemiAuto;
    countMem                : INT := 0;
END_VAR

{region "Corps d'exécution PRG_03 encapsulé"}
// 1. Arbitrage des Modes Machine
instModes(
    Enable                  := TRUE,
    Reset                   := BtnModeReset,
    PowerContactorEngaged   := PowerContactorEngaged,
    SelMode                 := SelMode,
    SelSyncEnable           := SelSyncEnable,
    InhibitM1Request        := InhibitM1Request,
    InhibitM2Request        := InhibitM2Request,
    SelHomingApproachEnable := SelHomingApproachEnable,
    EncoderFaultPresent     := EncoderFaultPresent,
    MachineHomed   := MachineHomed,
    JoystickWinchSelectRequest := SelJoystickWinch,
    SelMaintenanceZoneAccess := TglMaintenanceZoneAccess
);

Auth := instModes.Auth;

// 2. Séquenceur de Cycle Semi-Automatique
instCycleSemiAuto(
    Enable                  := (Auth.Mode = E_Mode.SEMI_AUTO),
    Reset                   := BtnCycleReset,
    PowerContactorEngaged   := PowerContactorEngaged,
    EncoderFaultPresent     := EncoderFaultPresent,
    Mode                    := Auth.Mode,
    CycleMotionPermit       := JoystickDeflected,
    DeadmanArmed            := DeadmanArmed,
    HeartbeatIhmOk          := HeartbeatIhmOk,
    StartCycle              := BtnStartCycle,
    AbortCycle              := BtnAbortCycle,
    SelTarget               := 1,
    SetDepthM               := -12.0,
    // SetOffsetM SUPPRIME (2026-09-22) : la VAR_INPUT n'existe plus sur FB_CycleSemiAuto
    // (retiree par le commit ffc811c1, audit CYCLE : « jamais utilisee »). Cet argument
    // mort bloquait la compilation g++ des entrees WINCH_INTEG, MAIN_GLOBAL et
    // PRG_03_Modes_Cycle (erreur « FB_CYCLESEMIAUTO has no member named SETOFFSETM »).
    // Preuve : TOOLS/TEST_AUTO_CI/RESULTS/H_TREUILS_BENNE/reports/WINCH_INTEG.txt.
    LimitLegalReached       := FALSE,
    LimitLegalDepthM        := -15.0,
    WinchSyncError          := FALSE,
    WinchSyncDeltaM         := 0.0,
    M1_CablePosM            := M1_CablePosM,
    M2_CablePosM            := M2_CablePosM,
    M1_MeasuredSpeedMps     := M1_SpeedMps,
    M2_MeasuredSpeedMps     := M2_SpeedMps,
    SpeedMismatchThresholdMps := 1.5,
    SpeedMismatchTimeout    := T#500ms,
    CableLimitM1AscentM     := 7.5,
    Translation_At_P1       := FALSE,
    Translation_At_Tremie   := TRUE,
    Translation_At_Maintenance := FALSE,
    Translation_Busy        := FALSE,
    Translation_Done        := TRUE,
    Benne_Busy              := FALSE,
    Benne_Done              := TRUE,
    Benne_IsOpen            := Benne_IsOpen,
    Benne_IsClosed          := Benne_IsClosed,
    Benne_IsRoughlyClosed   := Benne_IsRoughlyClosed,
    HomedM1                 := HomedM1,
    HomedM2                 := HomedM2,
    HomingRequest           := FALSE,
    SampleCount             := countMem
);

CycleStep     := instCycleSemiAuto.CycleStep;
CycleBusy     := instCycleSemiAuto.Lifecycle.Busy;
CycleDone     := instCycleSemiAuto.Lifecycle.Done;
CycleError    := instCycleSemiAuto.Fault.Error;
CycleStateStr := instCycleSemiAuto.CycleStateStr;

{endregion}
END_FUNCTION_BLOCK

(* ---- FB_TestHarness_PRG_04.st ---- *)
(*====================================================================
   FB_TestHarness_PRG_04 : Banc d'essai unitaire pour PRG_04_Treuils_Benne
   ==================================================================== *)

FUNCTION_BLOCK PUBLIC FB_TestHarness_PRG_04
VAR_IN_OUT
    BucketMech              : ST_fbBucket_State;
END_VAR

VAR_INPUT
    AcqData                : ST_AcquisitionInterPrg;
    ModesAuth               : ST_Modes_Autorisations;
    BtnWinchM1Up            : BOOL := FALSE;
    BtnWinchM1Down          : BOOL := FALSE;
    BtnWinchM2Up            : BOOL := FALSE;
    BtnWinchM2Down          : BOOL := FALSE;
    BtnWinchBothUp          : BOOL := FALSE;
    BtnWinchBothDown        : BOOL := FALSE;
    BucketBtnOpen           : BOOL := FALSE;
    BucketBtnClose          : BOOL := FALSE;
    PowerContactorEngaged   : BOOL := TRUE;
    M1_ContactorsReleased   : BOOL := TRUE;
    M2_ContactorsReleased   : BOOL := TRUE;
    M1_BrakeFeedbackOpen    : BOOL := TRUE;
    M2_BrakeFeedbackOpen    : BOOL := TRUE;
    M1_ThermalOk            : BOOL := TRUE;
    M2_ThermalOk            : BOOL := TRUE;
    BrakeThermalOk          : BOOL := TRUE;
    M1_TensionedCable       : BOOL := TRUE;
    M2_TensionedCable       : BOOL := TRUE;
    PhaseRotationOk         : BOOL := TRUE;
    TopPositionFreeDI       : BOOL := TRUE;
    TopHardStopLatched      : BOOL := FALSE;
    CfgTopEscalateDelay     : TIME := T#2s;
    BrakeForceAllowedM1     : BOOL := FALSE;
    FaultMachineResetIHM    : BOOL := FALSE;
    CfgCableLimitAscentM    : REAL := 7.5;
    CfgCableLimitDescentM1  : REAL := -30.0;
    CfgCableLimitDescentM2  : REAL := -30.0;
    WinchSlowdownDistanceM  : REAL := 1.0;
    WinchSlowdownMaxStep    : INT  := 1;
    SpeedStepTable          : ST_SpeedStepTable;
    BucketPersistConfig     : ST_fbBucket_Config;
END_VAR

VAR_OUTPUT
    Data                    : ST_WinchInterPrg;
END_VAR

VAR
    instWinchSync           : FB_WinchSync;
    instBucket              : FB_Bucket;
    instSafetyWinchM1       : FB_Safety_Winch;
    instSafetyWinchM2       : FB_Safety_Winch;
    instWinchM1             : FB_Winch;
    instWinchM2             : FB_Winch;
    ReqM1Winch              : ST_fbWinch_Req;
    ReqM2Winch              : ST_fbWinch_Req;
    M1WinchSensors          : ST_fbWinch_Sensors;
    M2WinchSensors          : ST_fbWinch_Sensors;
    M1WinchCfg              : ST_fbWinch_Cfg;
    M2WinchCfg              : ST_fbWinch_Cfg;
    M1LogicRunRequest       : BOOL;
    M1LogicReqAscent        : BOOL;
    M1LogicReqDescend       : BOOL;
    M1LogicRequestStepTgt   : INT;
    M1LogicRequestSpeedCmd_Pct : REAL;
    M2LogicRunRequest       : BOOL;
    M2LogicReqAscent        : BOOL;
    M2LogicReqDescend       : BOOL;
    M2LogicRequestStepTgt   : INT;
    M2LogicRequestSpeedCmd_Pct : REAL;
    SafeStopM1_Active       : BOOL;
    SafeStopM2_Active       : BOOL;
    EffectivePermitM1_Ascent : BOOL;
    EffectivePermitM1_Descend : BOOL;
    EffectivePermitM2_Ascent : BOOL;
    EffectivePermitM2_Descend : BOOL;
END_VAR

M1LogicReqAscent := BtnWinchM1Up OR (ModesAuth.JoystickWinchSelectArbitrated = 1 AND AcqData.Joystick.DeadmanArmed AND NOT AcqData.Joystick.AtNeutralXY AND (AcqData.Joystick.AxisY.Direction = 1));
M1LogicReqDescend := BtnWinchM1Down OR (ModesAuth.JoystickWinchSelectArbitrated = 1 AND AcqData.Joystick.DeadmanArmed AND NOT AcqData.Joystick.AtNeutralXY AND (AcqData.Joystick.AxisY.Direction = -1));
M1LogicRunRequest := M1LogicReqAscent OR M1LogicReqDescend;
M1LogicRequestStepTgt := SEL(M1LogicRunRequest, 0, 1);
M1LogicRequestSpeedCmd_Pct := SEL(M1LogicRunRequest, 0.0, 20.0);

M2LogicReqAscent := BtnWinchM2Up OR (ModesAuth.JoystickWinchSelectArbitrated = 2 AND AcqData.Joystick.DeadmanArmed AND NOT AcqData.Joystick.AtNeutralXY AND (AcqData.Joystick.AxisY.Direction = 1));
M2LogicReqDescend := BtnWinchM2Down OR (ModesAuth.JoystickWinchSelectArbitrated = 2 AND AcqData.Joystick.DeadmanArmed AND NOT AcqData.Joystick.AtNeutralXY AND (AcqData.Joystick.AxisY.Direction = -1));
M2LogicRunRequest := M2LogicReqAscent OR M2LogicReqDescend;
M2LogicRequestStepTgt := SEL(M2LogicRunRequest, 0, 1);
M2LogicRequestSpeedCmd_Pct := SEL(M2LogicRunRequest, 0.0, 20.0);

instSafetyWinchM1(
    Enable                  := (ModesAuth.Mode <> E_Mode.DISABLE) AND NOT ModesAuth.InhibitM1,
    Reset                   := FaultMachineResetIHM,
    Mode                    := ModesAuth.Mode,
    SyncEnable              := ModesAuth.SyncEnable,
    CrossCheckEnable        := ModesAuth.SyncEnable,
    ReqAscent               := M1LogicReqAscent,
    ReqDescend              := M1LogicReqDescend,
    MovementCommanded       := instWinchM1.RelayFwd OR instWinchM1.RelayRev,
    PowerContactorEngaged   := PowerContactorEngaged,
    JoystickOnline          := TRUE,
    JoystickOperational     := TRUE,
    HeartbeatIhmOk          := TRUE,
    EncoderAvailable        := AcqData.EncoderM1.Measurement.EncoderAvailable,
    ThermalFeedback         := NOT M1_ThermalOk,
    BrakeThermalFeedback    := NOT BrakeThermalOk,
    BypassOperatorComm      := TRUE,
    SlackCableDetected      := NOT M1_TensionedCable,
    PhaseRotationOk         := PhaseRotationOk,
    TopPositionSensor       := TopPositionFreeDI,
    FwdRevSpeedFeedbackOff  := M1_ContactorsReleased,
    BrakeFeedback           := M1_BrakeFeedbackOpen,
    JoystickYNeutral        := AcqData.Joystick.AtNeutralXY,
    CablePosM               := AcqData.EncoderM1.Measurement.CablePosM,
    CfgCableLimitDescentM   := CfgCableLimitDescentM1,
    TopLimitM               := CfgCableLimitAscentM,
    Homed                   := AcqData.EncoderM1.Homed,
    HomingSuspect           := AcqData.EncoderM1.HomingSuspect,
    MeasuredSpeedMps        := AcqData.EncoderM1.Measurement.Speed_Mps,
    MeasuredSpeedSignedMps  := AcqData.EncoderM1.Measurement.SignedSpeed_Mps,
    MeasuredSpeedValid      := AcqData.EncoderM1.Measurement.SpeedValid,
    SpeedBandMaxMps         := 2.0,
    BrakeForceAllowed       := BrakeForceAllowedM1,
    TopHardStopLatched      := TopHardStopLatched,
    CfgTopEscalateDelay     := CfgTopEscalateDelay
);

SafeStopM1_Active := instSafetyWinchM1.SafeStop;
EffectivePermitM1_Ascent := instSafetyWinchM1.AscentPermit AND NOT SafeStopM1_Active;
EffectivePermitM1_Descend := instSafetyWinchM1.DescendPermit AND NOT SafeStopM1_Active;

ReqM1Winch.RunRequest := M1LogicRunRequest;
ReqM1Winch.ReqAscent := M1LogicReqAscent;
ReqM1Winch.ReqDescend := M1LogicReqDescend;
ReqM1Winch.SpeedStepReq := M1LogicRequestStepTgt;
ReqM1Winch.MaxStepUp := 5;
ReqM1Winch.MaxStepDown := 3;

M1WinchSensors.CablePosM := AcqData.EncoderM1.Measurement.CablePosM;
M1WinchSensors.Homed := AcqData.EncoderM1.Homed;
M1WinchSensors.HomingSuspect := AcqData.EncoderM1.HomingSuspect;
M1WinchSensors.ContactorsAllOff := M1_ContactorsReleased;

M1WinchCfg.SpeedStepTable := SpeedStepTable;
M1WinchCfg.SlowdownDistanceBottom_M := WinchSlowdownDistanceM;
M1WinchCfg.SlowdownMaxStep := WinchSlowdownMaxStep;

instWinchM1(
    Enable                  := (ModesAuth.Mode <> E_Mode.DISABLE) AND NOT ModesAuth.InhibitM1,
    Reset                   := FaultMachineResetIHM,
    PowerContactorEngaged   := PowerContactorEngaged,
    SafeStop                := SafeStopM1_Active,
    DescendPermit           := EffectivePermitM1_Descend,
    AscentPermit            := EffectivePermitM1_Ascent,
    WinchRequest            := ReqM1Winch,
    Sensors                 := M1WinchSensors,
    Config                  := M1WinchCfg
);

Data.WinchM1FinalInterlockRequest.Enable := TRUE;
Data.WinchM1FinalInterlockRequest.Reset := FaultMachineResetIHM;
Data.WinchM1FinalInterlockRequest.PowerContactorEngaged := PowerContactorEngaged;
Data.WinchM1FinalInterlockRequest.SafeStop := SafeStopM1_Active;
Data.WinchM1FinalInterlockRequest.PowerCutOff := instSafetyWinchM1.PowerCutOff;
Data.WinchM1FinalInterlockRequest.AscentPermit := EffectivePermitM1_Ascent;
Data.WinchM1FinalInterlockRequest.DescendPermit := EffectivePermitM1_Descend;
Data.WinchM1FinalInterlockRequest.BrakeFeedback := M1_BrakeFeedbackOpen;
Data.WinchM1FinalInterlockRequest.FwdRevSpeedFeedbackOff := M1_ContactorsReleased;
Data.WinchM1FinalInterlockRequest.RequestedRelayFwd := M1LogicReqAscent AND NOT SafeStopM1_Active;
Data.WinchM1FinalInterlockRequest.RequestedRelayRev := M1LogicReqDescend AND NOT SafeStopM1_Active;
Data.WinchM1FinalInterlockRequest.RequestedContactor1 := instWinchM1.Contactor1;
Data.WinchM1FinalInterlockRequest.RequestedStep := instWinchM1.StepNumber;

Data.WinchM1Safety.SafeStop := SafeStopM1_Active;
Data.WinchM1Safety.PowerCutOff := instSafetyWinchM1.PowerCutOff;
Data.WinchM1Safety.Error := instSafetyWinchM1.Fault.Error;
Data.WinchM1Safety.ErrorId := instSafetyWinchM1.Fault.ErrorId;
Data.WinchM1Safety.LatchedId := instSafetyWinchM1.Fault.LatchedId;
Data.WinchM1Safety.ErrorMecaD := ((instSafetyWinchM1.Fault.ErrorId OR instSafetyWinchM1.Fault.LatchedId) AND 16#0800) <> 16#0000;
Data.WinchM1Safety.AscentPermit := EffectivePermitM1_Ascent;
Data.WinchM1Safety.DescendPermit := EffectivePermitM1_Descend;

Data.WinchM1State.RelayFwd := M1LogicReqAscent AND NOT SafeStopM1_Active;
Data.WinchM1State.RelayRev := M1LogicReqDescend AND NOT SafeStopM1_Active;
Data.WinchM1State.StepNumber := instWinchM1.StepNumber;

Data.M1LogicRequestSpeedCmd_Pct := M1LogicRequestSpeedCmd_Pct;

END_FUNCTION_BLOCK

(* ---- FB_TestHarness_PRG_05.st ---- *)
(* =======================================================================
   🧱 FB_TestHarness_PRG_05 : Banc d'essai unitaire pour PRG_05_Translation
   ───────────────────────────────────────────────────────────────
   🎯 Rôle : Isole PRG_05, consomme les bus de données de PRG_02 (Position,
             capteurs, joystick X), PRG_03 (Modes/Autorisations) et PRG_04 (Hauteur treuils),
             exécute FB_Translation et FB_Safety_Translation, et publie ST_TranslationInterPrg.
   ======================================================================= *)

FUNCTION_BLOCK PUBLIC FB_TestHarness_PRG_05
VAR_INPUT
    // === 📥 Bus d'Entrée issus de PRG_02 (Acquisition) ===
    AcqData                 : ST_AcquisitionInterPrg;

    // === 📥 Bus d'Entrée issus de PRG_03 (Modes) ===
    ModesAuth               : ST_Modes_Autorisations;

    // === 📥 Bus d'Entrée issus de PRG_04 (Treuils / Hauteur câble) ===
    WinchM1CablePosM        : REAL := 5.0;
    WinchM2CablePosM        : REAL := 5.0;

    // === 🛡️ Sécurités & Hardware Machine ===
    PowerContactorEngaged   : BOOL := TRUE;
    EmergencyChainClosed    : BOOL := TRUE;
    BrakeFeedbackOpen       : BOOL := FALSE;
    DriveOnline             : BOOL := TRUE;
    DriveOperational        : BOOL := TRUE;

    // === 🎛️ Commandes IHM Directes ===
    BtnReset                : BOOL := FALSE;
    BtnTranslationFwd       : BOOL := FALSE;
    BtnTranslationRev       : BOOL := FALSE;

    // === 🧩 Capteurs position M3 ===
    M3_PosTremie_DI         : BOOL := FALSE;
    M3_PosPV_DI             : BOOL := FALSE;
    M3_PosPVP2_DI           : BOOL := FALSE;
    M3_PosP1_DI             : BOOL := FALSE;
    M3_PosMaintenance_DI    : BOOL := FALSE;

    // === 🔒 Bypass IHM M3 (valeurs brutes : la garde de mode MAINT_N2 est appliquée par le harnais) ===
    BypassLimitSwitchIHM    : BOOL := FALSE;
    BypassGlobalIHM         : BOOL := FALSE;

    // === 🔌 Retour variateur M3 (injectable : au banc la fréquence réelle est nulle en permanence) ===
    DriveActualFreqHzOverride : REAL := 0.0;
END_VAR

VAR_OUTPUT
    // === 🚌 Bus Inter-PRG produit vers PRG_03/06/07 ===
    Data                    : ST_TranslationInterPrg;
END_VAR

VAR
    instTranslationM3       : FB_Translation;
    instSafetyTranslationM3 : FB_Safety_Translation;
    instPosDecoderM3        : FB_Translation_PositionDecoder;

    m3Cfg                   : ST_fbTranslation_Cfg;
    m3RunRequest            : BOOL;
    m3ReqTremie             : BOOL;
    m3ReqMaintenance        : BOOL;
    m3Direction             : INT;
    m3SpeedTgt              : REAL;
    m3HeightOk              : BOOL;
    initDone                : BOOL := FALSE;
    m3LimitSwitchTremieStable : BOOL;   // §0ter PRG_05 (guard REX MES 2026-09-04) : FdC latche, rebond capteur ne libere rien
    m3MaintN2               : BOOL;     // §1bis PRG_05 : mode MAINT_N2 arbitré (garde de consommation des bypass M3)
    m3PositionSensorTarget  : BOOL;     // §1 PRG_05 : cible d'arrêt publiée vers FB_Translation
    m3TargetCodeSel         : INT;      // §1 PRG_05 : code de cible mémorisé (1 = Trémie, 3 = P1)
    m3AtP1Stable            : BOOL;     // §0quater PRG_05 : jeton de point atteint P1
    m3AtTremieStable        : BOOL;     // §0quater PRG_05 : jeton de point atteint Trémie
    m3SensorsWordPrev       : BYTE;     // §0quater PRG_05 : mot capteurs du scan précédent
    m3SensorsWordChanged    : BOOL;     // §0quater PRG_05 : franchissement (mot capteurs changé)
END_VAR

{region "Corps d'exécution PRG_05 encapsulé"}
IF NOT initDone THEN
    m3Cfg.CfgRampAccelRate := 1000.0;
    m3Cfg.CfgRampDecelNormalRate := 1000.0;
    m3Cfg.CfgRampDecelFastRate := 2000.0;
    m3Cfg.DriveFreqScaleMaxHz := 50.0;
    initDone := TRUE;
END_IF;

// 0. Décodage position M3
instPosDecoderM3(
    SensorTremie      := M3_PosTremie_DI,
    SensorPV          := M3_PosPV_DI,
    SensorP2          := M3_PosPVP2_DI,
    SensorP1          := M3_PosP1_DI,
    SensorMaintenance := M3_PosMaintenance_DI
);

// 1. Interlock Hauteur Treuils
m3HeightOk := (WinchM1CablePosM >= 2.0) AND (WinchM2CablePosM >= 2.0);

// 2. Arbitrage Commande Translation
IF BtnTranslationFwd THEN
    m3ReqTremie      := TRUE;
    m3ReqMaintenance := FALSE;
    m3RunRequest     := TRUE;
    m3Direction      := 1;
    m3SpeedTgt       := 50.0;
ELSIF BtnTranslationRev THEN
    m3ReqTremie      := FALSE;
    m3ReqMaintenance := TRUE;
    m3RunRequest     := TRUE;
    m3Direction      := -1;
    m3SpeedTgt       := 50.0;
ELSIF AcqData.Joystick.DeadmanArmed AND (AcqData.Joystick.AxisX.Direction <> 0) AND m3HeightOk THEN
    m3ReqTremie      := (AcqData.Joystick.AxisX.Direction = 1);
    m3ReqMaintenance := (AcqData.Joystick.AxisX.Direction = -1);
    m3RunRequest     := TRUE;
    m3Direction      := AcqData.Joystick.AxisX.Direction;
    m3SpeedTgt       := ABS(AcqData.Joystick.AxisX.SpeedTgt);
ELSE
    m3ReqTremie      := FALSE;
    m3ReqMaintenance := FALSE;
    m3RunRequest     := FALSE;
    m3Direction      := 0;
    m3SpeedTgt       := 0.0;
END_IF;

// 2bis. Miroir réduit de PRG_05 §0quater, §1 et §1bis (T345/L1) — les trois faits touchés par le lot :
//   (a) jetons de point atteint Trémie/P1 armés sur le front du capteur propre et remis à zéro par
//       tout autre franchissement (miroir de PRG_05 §0quater) ;
//   (b) mémoire de cible : le code de cible n'est réécrit que tant qu'une demande est présente, la
//       cible publiée étant le jeton du point mémorisé (miroir de PRG_05 §1) ;
//   (c) garde de mode des bypass de fin de course : consommés uniquement en MAINT_N2 (miroir §1bis).
m3MaintN2 := (ModesAuth.Mode = E_Mode.MAINT_N2);

m3SensorsWordChanged := (instPosDecoderM3.SensorsWord <> m3SensorsWordPrev);
m3SensorsWordPrev := instPosDecoderM3.SensorsWord;

IF instPosDecoderM3.TranslationAtP1 THEN
    m3AtP1Stable := TRUE;
ELSIF instPosDecoderM3.TranslationAtTremie OR instPosDecoderM3.TranslationAtPV
      OR instPosDecoderM3.TranslationAtP2 OR instPosDecoderM3.TranslationAtMaintenance
      OR m3SensorsWordChanged THEN
    m3AtP1Stable := FALSE;
END_IF;

IF instPosDecoderM3.TranslationAtTremie THEN
    m3AtTremieStable := TRUE;
ELSIF instPosDecoderM3.TranslationAtPV OR instPosDecoderM3.TranslationAtP2
      OR instPosDecoderM3.TranslationAtP1 OR instPosDecoderM3.TranslationAtMaintenance
      OR m3SensorsWordChanged THEN
    m3AtTremieStable := FALSE;
END_IF;

IF m3ReqTremie THEN
    m3TargetCodeSel := 1;
ELSIF m3ReqMaintenance THEN
    m3TargetCodeSel := 3;
END_IF;

CASE m3TargetCodeSel OF
    1: m3PositionSensorTarget := m3AtTremieStable;
    3: m3PositionSensorTarget := m3AtP1Stable;
ELSE
    m3PositionSensorTarget := FALSE;
END_CASE;

// 3. Sécurité Translation M3
instSafetyTranslationM3(
    Enable                  := (ModesAuth.Mode <> E_Mode.DISABLE),
    Reset                   := BtnReset,
    PowerContactorEngaged   := PowerContactorEngaged,
    Mode                    := ModesAuth.Mode,
    JoystickOnline          := TRUE,
    JoystickOperational     := TRUE,
    HeartbeatIhmOk          := TRUE,
    PhaseRotationOk         := TRUE,
    BrakeThermalFeedback    := FALSE,
    DriveOnline             := DriveOnline,
    DriveOperational        := DriveOperational,
    DriveStatusWord         := 16#0000,
    DriveActualFreqHz       := DriveActualFreqHzOverride,
    BrakeFeedback           := BrakeFeedbackOpen,
    BrakeCmd                := FALSE,
    RunRequest              := m3RunRequest,
    ReqTremie               := m3ReqTremie,
    ReqMaintenance          := m3ReqMaintenance,
    LimitSwitchTremie       := instPosDecoderM3.LimitSwitchTremie,
    LimitSwitchMaintenance  := instPosDecoderM3.LimitSwitchMaintenance,
    SensorWordIncoherent    := instPosDecoderM3.Incoherent,
    BypassLimitSwitch       := m3MaintN2 AND (BypassLimitSwitchIHM OR BypassGlobalIHM)
);

Data.TranslationSafety.SafeStop    := instSafetyTranslationM3.SafeStop;
Data.TranslationSafety.PowerCutOff := instSafetyTranslationM3.PowerCutOff;

// 4. Pilotage M3
instTranslationM3(
    Enable                     := (ModesAuth.Mode <> E_Mode.DISABLE),
    Reset                      := BtnReset,
    PowerContactorEngaged      := PowerContactorEngaged,
    Mode                       := ModesAuth.Mode,
    RunRequest                 := m3RunRequest,
    SafeStop                   := Data.TranslationSafety.SafeStop,
    ReqTremie                  := m3ReqTremie,
    ReqMaintenance             := m3ReqMaintenance,
    SpeedTgt_Pct               := m3SpeedTgt,
    PositionSensorTarget       := m3PositionSensorTarget,
    SlowdownSensorTremie       := instPosDecoderM3.TranslationPosPV,
    SlowdownSensorMaintenance  := instPosDecoderM3.TranslationPosP1,
    SlowdownSensorP1           := instPosDecoderM3.TranslationPosP2,
    LimitSwitchTremie          := instPosDecoderM3.LimitSwitchTremie,
    LimitSwitchMaintenance     := instPosDecoderM3.LimitSwitchMaintenance,
    EffectivePermitM3_Tremie   := instSafetyTranslationM3.TremieLimitClear,
    EffectivePermitM3_Maintenance := instSafetyTranslationM3.MaintenanceLimitClear,
    DriveStatusWord            := 16#0081,
    DriveActualFreqHz          := DriveActualFreqHzOverride,
    BrakeFeedback              := BrakeFeedbackOpen,
    BypassLimitSwitch          := m3MaintN2 AND (BypassLimitSwitchIHM OR BypassGlobalIHM),
    Cfg                        := m3Cfg
);

// 5. Remplissage Bus Sortie Data
Data.TranslationFinalInterlockRequest.Enable                    := instTranslationM3.Enable;
Data.TranslationFinalInterlockRequest.Reset                     := BtnReset;
Data.TranslationFinalInterlockRequest.PowerContactorEngaged     := PowerContactorEngaged;
Data.TranslationFinalInterlockRequest.SafeStop                  := Data.TranslationSafety.SafeStop;
Data.TranslationFinalInterlockRequest.PowerCutOff               := Data.TranslationSafety.PowerCutOff;
Data.TranslationFinalInterlockRequest.BrakeReleaseRequest       := instTranslationM3.BrakeReleaseRequest;
Data.TranslationFinalInterlockRequest.RequestedDriveControlWord := instTranslationM3.RequestedDriveControlWord;
Data.TranslationFinalInterlockRequest.RequestedDriveFreqHz      := instTranslationM3.RequestedDriveFreqHz;

// §0ter PRG_05 : bistable FdC Tremie LATCHE. Un rebond capteur (mot 11111 <-> 01111)
// ne libere RIEN. Perte de la butee UNIQUEMENT sur commande sens inverse (Maintenance).
IF instPosDecoderM3.LimitSwitchTremie THEN
    m3LimitSwitchTremieStable := TRUE;
ELSIF (m3Direction = -1) THEN
    m3LimitSwitchTremieStable := FALSE;
END_IF;
Data.TranslationState.LimitSwitchTremie := m3LimitSwitchTremieStable;

Data.TranslationState.ActiveTremie := (m3Direction = 1);
Data.TranslationState.ActiveMaintenance := (m3Direction = -1);
Data.TranslationState.SpeedCmd_Pct                             := m3SpeedTgt;
Data.TranslationState.Busy                                     := (instTranslationM3.RequestedDriveControlWord <> 0);
Data.TranslationState.Ready                                    := instTranslationM3.Ready;
// Publication des faits observés par la porte de cycle (mêmes champs que PRG_05) :
// la cible qualifiée de l'axe et son défaut propre.
Data.TranslationDone                                           := instTranslationM3.TargetReached;
Data.TranslationState.Error                                    := instTranslationM3.Fault.Error;
{endregion}
END_FUNCTION_BLOCK

(* ---- FB_TestHarness_PRG_06.st ---- *)
(* =======================================================================
   🧱 FB_TestHarness_PRG_06 : Banc d'essai unitaire pour PRG_06_Outputs
   ───────────────────────────────────────────────────────────────
   🎯 Rôle : Isole PRG_06_Outputs, consomme les bus de données de
             PRG_04 (ST_WinchInterPrg) et PRG_05 (ST_TranslationInterPrg),
             exécute les barrières finales FB_WinchOutputInterlock (M1, M2)
             et FB_TranslationOutputInterlock (M3), et publie ST_OutputsInterPrg.
   ======================================================================= *)

FUNCTION_BLOCK PUBLIC FB_TestHarness_PRG_06
VAR_INPUT
    // === 📥 Bus d'Entrée issus de PRG_04 (Treuils M1/M2) ===
    WinchData                        : ST_WinchInterPrg;

    // === 📥 Bus d'Entrée issus de PRG_05 (Translation M3) ===
    TranslationData                  : ST_TranslationInterPrg;

    // === 🛡️ Entrées Supervision / Reset ===
    FaultReset                       : BOOL := FALSE;
    TopPositionFreeDI                : BOOL := TRUE;
    BypassTopLimitSwitch             : BOOL := FALSE;
    BypassM1TopLimitSwitch           : BOOL := FALSE;
    BypassM2TopLimitSwitch           : BOOL := FALSE;
END_VAR

VAR_OUTPUT
    // === 🚌 Bus Inter-PRG produit vers PRG_02/SimBench ===
    Data                             : ST_OutputsInterPrg;

    // Diagnostic
    M1InterlockEnable                : BOOL;
    M2InterlockEnable                : BOOL;
    M3InterlockEnable                : BOOL;
END_VAR

VAR
    instWinchOutputInterlockM1       : FB_WinchOutputInterlock;
    instWinchOutputInterlockM2       : FB_WinchOutputInterlock;
    instTranslationOutputInterlockM3 : FB_TranslationOutputInterlock;
    TopHardStopClearTimer            : TON;
    TopBypassM1                      : BOOL;
    TopBypassM2                      : BOOL;
    TopBypassAll                     : BOOL;
    M1_TopHardStopBlocked            : BOOL;
    M2_TopHardStopBlocked            : BOOL;
END_VAR

VAR RETAIN
    M1M2_TopHardStopLatched          : BOOL := FALSE;
END_VAR

{region "Corps d'exécution PRG_06 encapsulé"}
// 1. Barrière M1
M1InterlockEnable := WinchData.WinchM1FinalInterlockRequest.Enable
                     AND NOT WinchData.WinchM1FinalInterlockRequest.PowerCutOff;
TopBypassM1 := BypassTopLimitSwitch OR BypassM1TopLimitSwitch;
TopBypassM2 := BypassTopLimitSwitch OR BypassM2TopLimitSwitch;
TopBypassAll := BypassTopLimitSwitch OR (TopBypassM1 AND TopBypassM2);
IF NOT TopPositionFreeDI AND NOT TopBypassAll THEN
    M1M2_TopHardStopLatched := TRUE;
END_IF;
TopHardStopClearTimer(
    IN := M1M2_TopHardStopLatched
          AND TopPositionFreeDI
          AND (WinchData.WinchM1FinalInterlockRequest.RequestedRelayRev
               OR WinchData.WinchM2FinalInterlockRequest.RequestedRelayRev)
          AND NOT WinchData.WinchM1FinalInterlockRequest.RequestedRelayFwd
          AND NOT WinchData.WinchM2FinalInterlockRequest.RequestedRelayFwd,
    PT := T#3s
);
IF TopHardStopClearTimer.Q OR (FaultReset AND (TopPositionFreeDI OR TopBypassAll)) THEN
    M1M2_TopHardStopLatched := FALSE;
END_IF;
M1_TopHardStopBlocked := (NOT TopPositionFreeDI OR M1M2_TopHardStopLatched) AND NOT TopBypassM1;
M2_TopHardStopBlocked := (NOT TopPositionFreeDI OR M1M2_TopHardStopLatched) AND NOT TopBypassM2;

instWinchOutputInterlockM1(
    Enable                     := M1InterlockEnable,
    Reset                      := FaultReset,
    PowerContactorEngaged      := WinchData.WinchM1FinalInterlockRequest.PowerContactorEngaged,
    SafeStop                   := WinchData.WinchM1FinalInterlockRequest.SafeStop,
    AscentPermit               := WinchData.WinchM1FinalInterlockRequest.AscentPermit AND NOT M1_TopHardStopBlocked,
    DescendPermit              := WinchData.WinchM1FinalInterlockRequest.DescendPermit,
    BrakeFeedback              := WinchData.WinchM1FinalInterlockRequest.BrakeFeedback,
    FwdRevSpeedFeedbackOff     := WinchData.WinchM1FinalInterlockRequest.FwdRevSpeedFeedbackOff,
    RequestedRelayFwd          := WinchData.WinchM1FinalInterlockRequest.RequestedRelayFwd,
    RequestedRelayRev          := WinchData.WinchM1FinalInterlockRequest.RequestedRelayRev,
    RequestedContactor1        := WinchData.WinchM1FinalInterlockRequest.RequestedContactor1,
    RequestedContactor2        := WinchData.WinchM1FinalInterlockRequest.RequestedContactor2,
    RequestedContactor3        := WinchData.WinchM1FinalInterlockRequest.RequestedContactor3,
    RequestedContactor4        := WinchData.WinchM1FinalInterlockRequest.RequestedContactor4,
    RequestedStep              := WinchData.WinchM1FinalInterlockRequest.RequestedStep
);

Data.M1RelayFwd        := instWinchOutputInterlockM1.RelayFwd;
Data.M1RelayRev        := instWinchOutputInterlockM1.RelayRev;
Data.M1SpeedContactor1 := instWinchOutputInterlockM1.Contactor1;
Data.M1SpeedContactor2 := instWinchOutputInterlockM1.Contactor2;
Data.M1SpeedContactor3 := instWinchOutputInterlockM1.Contactor3;
Data.M1SpeedContactor4 := instWinchOutputInterlockM1.Contactor4;
Data.M1BrakeCmd        := Data.M1RelayFwd OR Data.M1RelayRev;

// 2. Barrière M2
M2InterlockEnable := WinchData.WinchM2FinalInterlockRequest.Enable
                     AND NOT WinchData.WinchM2FinalInterlockRequest.PowerCutOff;

instWinchOutputInterlockM2(
    Enable                     := M2InterlockEnable,
    Reset                      := FaultReset,
    PowerContactorEngaged      := WinchData.WinchM2FinalInterlockRequest.PowerContactorEngaged,
    SafeStop                   := WinchData.WinchM2FinalInterlockRequest.SafeStop,
    AscentPermit               := WinchData.WinchM2FinalInterlockRequest.AscentPermit AND NOT M2_TopHardStopBlocked,
    DescendPermit              := WinchData.WinchM2FinalInterlockRequest.DescendPermit,
    BrakeFeedback              := WinchData.WinchM2FinalInterlockRequest.BrakeFeedback,
    FwdRevSpeedFeedbackOff     := WinchData.WinchM2FinalInterlockRequest.FwdRevSpeedFeedbackOff,
    RequestedRelayFwd          := WinchData.WinchM2FinalInterlockRequest.RequestedRelayFwd,
    RequestedRelayRev          := WinchData.WinchM2FinalInterlockRequest.RequestedRelayRev,
    RequestedContactor1        := WinchData.WinchM2FinalInterlockRequest.RequestedContactor1,
    RequestedContactor2        := WinchData.WinchM2FinalInterlockRequest.RequestedContactor2,
    RequestedContactor3        := WinchData.WinchM2FinalInterlockRequest.RequestedContactor3,
    RequestedContactor4        := WinchData.WinchM2FinalInterlockRequest.RequestedContactor4,
    RequestedStep              := WinchData.WinchM2FinalInterlockRequest.RequestedStep
);

Data.M2RelayFwd        := instWinchOutputInterlockM2.RelayFwd;
Data.M2RelayRev        := instWinchOutputInterlockM2.RelayRev;
Data.M2SpeedContactor1 := instWinchOutputInterlockM2.Contactor1;
Data.M2SpeedContactor2 := instWinchOutputInterlockM2.Contactor2;
Data.M2SpeedContactor3 := instWinchOutputInterlockM2.Contactor3;
Data.M2SpeedContactor4 := instWinchOutputInterlockM2.Contactor4;
Data.M2BrakeCmd        := Data.M2RelayFwd OR Data.M2RelayRev;

// 3. Barrière M3
M3InterlockEnable := TranslationData.TranslationFinalInterlockRequest.Enable
                     AND NOT TranslationData.TranslationFinalInterlockRequest.PowerCutOff;

instTranslationOutputInterlockM3(
    Enable                     := M3InterlockEnable,
    Reset                      := FaultReset,
    PowerContactorEngaged      := TranslationData.TranslationFinalInterlockRequest.PowerContactorEngaged,
    SafeStop                   := TranslationData.TranslationFinalInterlockRequest.SafeStop,
    BrakeCommandOpenConfirmed  := TranslationData.TranslationFinalInterlockRequest.BrakeCommandOpenConfirmed,
    BrakeReleaseRequest        := TranslationData.TranslationFinalInterlockRequest.BrakeReleaseRequest,
    RequestedDriveControlWord  := TranslationData.TranslationFinalInterlockRequest.RequestedDriveControlWord,
    RequestedDriveFreqHz       := TranslationData.TranslationFinalInterlockRequest.RequestedDriveFreqHz
);

Data.TranslationBrakeCmd := instTranslationOutputInterlockM3.BrakeCmd;
Data.TopHardStopLatched := M1M2_TopHardStopLatched;

{endregion}
END_FUNCTION_BLOCK

(* ---- FB_TestHarness_PRG_07.st ---- *)
(* =======================================================================
   🧱 FB_TestHarness_PRG_07 : Banc d'essai unitaire pour PRG_07_Supervision
   ───────────────────────────────────────────────────────────────
   🎯 Rôle : Isole PRG_07_Supervision, consomme les bus de données
             de PRG_02 (Joystick/E-S), PRG_03 (Modes/Cycle), PRG_04 (Treuils/Benne)
             et PRG_05 (Translation), exécute le formateur de bandeau
             FB_Hmi_BannerFormatter et publie le bandeau IHM ST_HmiBanner.
   ======================================================================= *)

FUNCTION_BLOCK PUBLIC FB_TestHarness_PRG_07
VAR_INPUT
    // === 📥 Bus d'Entrée issus de PRG_02 (Acquisition) ===
    AcqData                 : ST_AcquisitionInterPrg;

    // === 📥 Bus d'Entrée issus de PRG_03 (Modes & Cycle) ===
    ModesAuth               : ST_Modes_Autorisations;

    // === 📥 Bus d'Entrée issus de PRG_04 (Treuils & Benne) ===
    WinchData               : ST_WinchInterPrg;

    // === 📥 Bus d'Entrée issus de PRG_05 (Translation M3) ===
    TranslationData         : ST_TranslationInterPrg;

    // === 🛡️ État public de la chaîne AU (miroir de PRG_06_Outputs.EmergencyState) ===
    // Step : 0 = IDLE ; ContactorOk : contacteur de puissance confirmé engagé.
    EmergencyState          : ST_Safety_Emergency_State;

    // === 🛡️ Hardware & Sécurité Machine ===
    EmergencyChainClosed    : BOOL := TRUE;
    PowerContactorEngaged   : BOOL := TRUE;
    PowerCutOffActive       : BOOL := FALSE;
    BtnResetMachine         : BOOL := FALSE;
    TopHardStopLatched      : BOOL := FALSE;
    TopPositionSensorActive : BOOL := FALSE;
    Network                 : ST_NetworkDiagHMI;
END_VAR

VAR_OUTPUT
    // === 🖥️ Bandeau IHM Produit ===
    Banner                  : ST_HmiBanner;
    FaultMachineReset_IHM   : BOOL;
    AnyFaultActive          : BOOL;

    // === 🚨 Campagnes d'acquittement automatique borné (miroir PRG_07 §1c-1) ===
    BootAckPulse            : BOOL; // Impulsion émise par la campagne de démarrage à froid
    RearmAckPulse           : BOOL; // Impulsion émise par la campagne de réarmement AU
    BootAckFinished         : BOOL; // Campagne de démarrage à froid terminée (arrêt définitif)
END_VAR

VAR
    instHmiBannerFormatter  : FB_Hmi_BannerFormatter;

    // === 🚨 Campagnes d'acquittement automatique borné (miroir PRG_07_Supervision §1c-1) ===
    // États LOCAUX NON RETAIN, comme dans le PROGRAM : une campagne de démarrage à froid
    // ne peut pas se relancer sans un nouveau démarrage à froid.
    BootInputTransientDone : BOOL;   // Transitoire d'E/S terminé (5 modules RUNNING)
    BootWindowTimer        : TON;    // Fenêtre de démarrage à froid (borne la campagne)
    BootSettleTimer        : TON;    // Tempo de stabilisation après le transitoire d'E/S
    BootAckWindowOpen      : BOOL;   // Fenêtre de démarrage à froid encore ouverte
    BootAckStart           : BOOL;   // Campagne de démarrage à froid à démarrer
    BootCampaignLastPulse  : BOOL;   // Dernière impulsion de la campagne de démarrage à froid
    BootCampaignEnded      : BOOL;   // Campagne de démarrage à froid close
    RearmSeqRunning        : BOOL;   // Une séquence d'armement AU est en cours (Step <> 0)
    RearmSeqStartEdge      : R_TRIG; // Front de démarrage d'une séquence d'armement
    RearmSeqSeen           : BOOL;   // Une séquence d'armement a démarré (geste opérateur)
    RearmGestureTimer      : TON;    // Durée de vie du geste d'armement (anti-mémoire périmée)
    ContactorOkEdge        : R_TRIG; // Front montant du contacteur de puissance
    RearmAckStart          : BOOL;   // Campagne de réarmement AU à démarrer
    RearmCampaignLastPulse : BOOL;   // Dernière impulsion de la campagne de réarmement
    AckCampaignActive      : BOOL;   // Une campagne d'acquittement automatique est en cours
    AckCampaignIsBoot      : BOOL;   // La campagne en cours est celle du démarrage à froid
    AckPulseSpacing        : TON;    // Intervalle entre deux impulsions d'une campagne
    AckPulseCount          : USINT;  // Impulsions déjà émises par la campagne en cours
    AckPulseRoom           : BOOL;   // La campagne en cours a encore le droit d'impulsion
    AckPulseDue            : BOOL;   // Échéance d'impulsion atteinte
    AckCampaignPulsing     : BOOL;   // La campagne en cours a le droit d'émettre maintenant
    AckPulseAllowed        : BOOL;   // Acquittement autorisé (fin du transitoire d'E/S en boot)
    AckPulse               : BOOL;   // Impulsion d'acquittement de la campagne en cours
END_VAR

VAR CONSTANT
    // === 🚨 ACQUITTEMENT AUTOMATIQUE — BORNES DE CAMPAGNE (mêmes valeurs que PRG_07) ===
    CST_AckBootWindow   : TIME  := T#30s;
    CST_AckBootSettle   : TIME  := T#3s;
    CST_AckPulseSpacing : TIME  := T#1s;
    CST_AckPulseMax     : USINT := 3;
    CST_RearmGestureTtl : TIME  := T#10s;  // Durée de vie d'un geste non confirmé (identique à PRG_07)
END_VAR

{region "Corps d'exécution PRG_07 encapsulé"}
// 1. Gestion Reset Machine
// §1c-1. Campagnes d'acquittement AUTOMATIQUE BORNE — miroir strict de PRG_07_Supervision.
// (a) DÉMARRAGE À FROID : aucune impulsion tant que le transitoire d'E/S n'est pas terminé,
//     puis temps de stabilisation ; la fenêtre de démarrage borne la campagne.
// (b) RÉARMEMENT AU : une séquence d'armement doit avoir réellement démarré (front de Step)
//     avant le front du contacteur de puissance — le seul front du contacteur ne suffit jamais.
BootInputTransientDone := NOT AcqData.InputModules.Fault;
BootWindowTimer(IN := TRUE, PT := CST_AckBootWindow);
BootAckWindowOpen := NOT BootWindowTimer.Q;
BootSettleTimer(IN := BootInputTransientDone AND NOT BootAckFinished, PT := CST_AckBootSettle);
BootAckStart := BootSettleTimer.Q AND NOT BootAckFinished AND BootAckWindowOpen;

RearmSeqRunning := (EmergencyState.Step <> 0);
RearmSeqStartEdge(CLK := RearmSeqRunning);
IF RearmSeqStartEdge.Q THEN
    RearmSeqSeen := TRUE;
END_IF;
ContactorOkEdge(CLK := EmergencyState.ContactorOk);
RearmAckStart := ContactorOkEdge.Q AND RearmSeqSeen;
IF RearmAckStart THEN
    RearmSeqSeen := FALSE; // geste consommé : une nouvelle campagne exige un nouveau geste
END_IF;
// Durée de vie du geste : un armement ÉCHOUÉ ne doit pas laisser une mémoire consommable plus tard
// par un front du contacteur purement machine (relâchement d'un AU, maintien repris).
RearmGestureTimer(IN := RearmSeqSeen AND NOT ContactorOkEdge.Q, PT := CST_RearmGestureTtl);
IF RearmGestureTimer.Q THEN RearmSeqSeen := FALSE; END_IF; // geste périmé : nouveau geste requis

IF (BootAckStart OR RearmAckStart) AND NOT AckCampaignActive THEN
    AckCampaignActive := TRUE;
    AckCampaignIsBoot := BootAckStart;
    AckPulseCount     := 0;
END_IF;

AckPulseSpacing(IN := AckCampaignActive AND NOT AckPulseSpacing.Q, PT := CST_AckPulseSpacing);
AckPulseAllowed := TRUE;
IF AckCampaignIsBoot THEN
    AckPulseAllowed := BootInputTransientDone;
END_IF;
AckPulseRoom       := AckPulseCount < CST_AckPulseMax;
AckPulseDue        := (AckPulseCount = 0) OR AckPulseSpacing.Q;
AckCampaignPulsing := AckCampaignActive AND AckPulseAllowed AND AckPulseRoom;
AckPulse           := AckCampaignPulsing AND AckPulseDue;
IF AckPulse THEN
    AckPulseCount := AckPulseCount + 1;
END_IF;
BootAckPulse  := AckPulse AND AckCampaignIsBoot;
RearmAckPulse := AckPulse AND NOT AckCampaignIsBoot;

BootCampaignLastPulse := AckCampaignActive AND AckCampaignIsBoot AND (AckPulseCount >= CST_AckPulseMax);
BootCampaignEnded     := (NOT BootAckWindowOpen) OR BootCampaignLastPulse;
IF NOT BootAckFinished AND BootCampaignEnded THEN
    BootAckFinished := TRUE;
    IF AckCampaignIsBoot THEN
        AckCampaignActive := FALSE;
    END_IF;
END_IF;

RearmCampaignLastPulse := AckCampaignActive AND (NOT AckCampaignIsBoot) AND (AckPulseCount >= CST_AckPulseMax);
IF RearmCampaignLastPulse THEN
    AckCampaignActive := FALSE;
END_IF;

// §1c-2. Porte unique d'acquittement machine
FaultMachineReset_IHM := BtnResetMachine OR BootAckPulse OR RearmAckPulse;

// 2. Formatage Bandeau IHM
instHmiBannerFormatter(
    Enable                := TRUE,
    SimulationModeActive  := FALSE,
    CurrentMode           := ModesAuth.Mode,
    BothAxesCoupled       := (ModesAuth.JoystickWinchSelectArbitrated = 0),
    WinchSelected         := ModesAuth.JoystickWinchSelectArbitrated,
    CycleStep             := E_AutoCycleStep.AX0_REPOS,
    CycleStateStr         := 'X0_PREPARATION',
    CycleErrorId          := 16#0000,
    CycleStepAtError      := E_AutoCycleStep.AX0_REPOS,
    MachineHomingStep     := AcqData.MachineHoming.Step,
    MachineHomingInstruction := AcqData.MachineHoming.Instruction,
    MachineHomingFailed   := AcqData.MachineHoming.Failed,
    MachineHomingLoss     := AcqData.MachineHoming.HomingLoss,
    TopHardStopLatched    := TopHardStopLatched,
    TopPositionSensorActive := TopPositionSensorActive,
    WinchM1Error          := WinchData.WinchM1State.Error OR WinchData.WinchM1State.FaultLatched OR WinchData.WinchM1State.FinalInterlockError,
    WinchM2Error          := WinchData.WinchM2State.Error OR WinchData.WinchM2State.FaultLatched OR WinchData.WinchM2State.FinalInterlockError,
    SyncFaultLatched      := WinchData.SyncState.FaultLatched,
    BucketFaultLatched    := WinchData.BucketState.FaultLatched,
    EncoderM1Fault        := AcqData.EncoderM1.Fault.Error OR AcqData.EncoderM1.Fault.Latched,
    EncoderM2Fault        := AcqData.EncoderM2.Fault.Error OR AcqData.EncoderM2.Fault.Latched,
    JoystickLatchedFault  := AcqData.Joystick.Fault.Latched,

    BypassGlobalActive    := FALSE,
    BypassWinchM1Active   := FALSE,
    BypassWinchM2Active   := FALSE,
    BypassTranslation     := FALSE,
    BypassSyncActive      := FALSE,
    SyncDegradedActive    := FALSE,
    LegalLimitReached     := FALSE,
    EmergencyChainClosed  := EmergencyChainClosed,
    PowerContactorEngaged := PowerContactorEngaged,
    PowerCutOffActiveAny  := PowerCutOffActive,
    SafeStopActive        := WinchData.WinchM1Safety.SafeStop OR WinchData.WinchM2Safety.SafeStop,
    DescendPermit         := WinchData.WinchM1Safety.DescendPermit AND WinchData.WinchM2Safety.DescendPermit,
    AscentPermit          := WinchData.WinchM1Safety.AscentPermit AND WinchData.WinchM2Safety.AscentPermit,
    BucketIsOpen          := WinchData.BucketState.MechState.IsOpen,
    BucketIsClosed        := WinchData.BucketState.MechState.IsClosed,
    DiveActive            := FALSE,
    TopLimitReached       := WinchData.WinchM1Safety.CableLimitAscent OR WinchData.WinchM2Safety.CableLimitAscent,
    WinchBothMotionDirection := 0,
    M1LogicRequestDirection     := 0,
    M2LogicRequestDirection     := 0,
    CycleRequestDirection       := 0,
    DeadmanArmed          := AcqData.Joystick.DeadmanArmed,
    JoystickAtNeutral     := AcqData.Joystick.AtNeutralXY,
    CycleAutoBusy         := FALSE,
    WinchM1Safety         := WinchData.WinchM1Safety,
    WinchM2Safety         := WinchData.WinchM2Safety,
    TranslationSafety     := TranslationData.TranslationSafety,
    BucketErrorId         := 16#0000,
    SyncErrorId           := 16#0000,
    DiveErrorId           := 16#0000,
    ExtractionErrorId     := 16#0000,
    EmergencyErrorId      := 16#0000,
    RedundancyTestFailed  := FALSE,
    EmergencyArmingFailed := FALSE,
    AlarmHoldTime         := T#1s,
    Network               := Network
);

Banner := instHmiBannerFormatter.Banner;
AnyFaultActive := AcqData.InputModules.Fault
                  OR AcqData.MachineHoming.Failed
                  OR AcqData.MachineHoming.HomingLoss
                  OR AcqData.EncoderM1.Fault.Error
                  OR AcqData.EncoderM1.Fault.Latched
                  OR AcqData.EncoderM2.Fault.Error
                  OR AcqData.EncoderM2.Fault.Latched
                  OR AcqData.Joystick.Fault.Latched
                  OR WinchData.WinchM1Safety.Error
                  OR WinchData.WinchM1Safety.ErrorOverspeed
                  OR (WinchData.WinchM1Safety.LatchedId <> 16#0000)
                  OR WinchData.WinchM1State.Error
                  OR WinchData.WinchM1State.FaultLatched
                  OR WinchData.WinchM1State.FinalInterlockError
                  OR WinchData.WinchM2Safety.Error
                  OR WinchData.WinchM2Safety.ErrorOverspeed
                  OR (WinchData.WinchM2Safety.LatchedId <> 16#0000)
                  OR WinchData.WinchM2State.Error
                  OR WinchData.WinchM2State.FaultLatched
                  OR WinchData.WinchM2State.FinalInterlockError
                  OR TranslationData.TranslationSafety.Error
                  OR (TranslationData.TranslationSafety.LatchedId <> 16#0000)
                  OR TranslationData.TranslationState.Error
                  OR TranslationData.TranslationState.FinalInterlockError
                  OR WinchData.SyncState.Error
                  OR WinchData.SyncState.FaultLatched
                  OR WinchData.BucketState.Error
                  OR WinchData.BucketState.FaultLatched;
{endregion}
END_FUNCTION_BLOCK
